// TIA Portal V18 export
// export: Created 2026-11-25T00:00:00.0000000Z, ExportSetting WithDefaults
Screen "Alarms"  800x480, Number=3
  ScreenLayer 
    TextField "Title" at 8,8 size 600x28  Text="Alarms"
    TextField "Note" at 8,50 size 780x120  Text="Station alarms are Program_Alarm instances in the CPU (FB_StationAlarms): safety circuit open, drive not ready, clamp time-out, tare failed, reject waiting, rig check. Fault code now:"
    IOField "VFaultCode" at 8,180 size 140x30  FormatPattern=s999999, Mode=Output
      ProcessValue := FaultCode
    TextField "LCall" at 8,220 size 420x30  Text="Operator called"
    IOField "VCall" at 440,220 size 140x30  FormatPattern=9, Mode=Output
      ProcessValue := CallOperator
    Button "NavStation" at 8,424 size 188x48  TextOff="Station", TextOn="Station"
      on Click: ActivateScreen(Screen name := Station)
    Button "NavMeasurement" at 204,424 size 188x48  TextOff="Measurement", TextOn="Measurement"
      on Click: ActivateScreen(Screen name := Measurement)
    Button "NavAlarms" at 400,424 size 188x48  TextOff="Alarms", TextOn="Alarms"
      on Click: ActivateScreen(Screen name := Alarms)
    Button "NavSetup" at 596,424 size 188x48  TextOff="Setup", TextOn="Setup"
      on Click: ActivateScreen(Screen name := Setup)
